// TIA Portal V19 export
DATA_BLOCK "Valves Data"   // DB3
{ S7_Optimized_Access := 'FALSE'; DB_Accessible_From_OPC_UA := 'FALSE' }
// stored: DBAccessibleFromOPCUA false
   VAR RETAIN
      "A/M" : Struct
         R1 : Bool;
         R2 : Bool;
         R3 : Bool;
         R4 : Bool;
         R5 : Bool;
         R6 : Bool;
         R7 : Bool;
         R8 : Bool;
         R9 : Bool;
         R10 : Bool;
         R11 : Bool;
         R12 : Bool;
         R13 : Bool;
         R14 : Bool;
         R15 : Bool;
         R16 : Bool;
         R17 : Bool;
         R18 : Bool;
      END_STRUCT;
      SEMI_AUTO : Struct
         R1 : Bool;
         R2 : Bool;
         R3 : Bool;
         R4 : Bool;
         R5 : Bool;
         R6 : Bool;
         R7 : Bool;
         R8 : Bool;
         R9 : Bool;
         R10 : Bool;
         R11 : Bool;
         R12 : Bool;
         R13 : Bool;
         R14 : Bool;
         R15 : Bool;
         R16 : Bool;
         R17 : Bool;
         R18 : Bool;
      END_STRUCT;
      R1_XV01 : Struct
         MCMD : Bool;
         CMD : Bool;
         RESET : Bool;
         MON_TIME : Time := T#5S;
         STATUS : Int;
         FAULTY : Bool;
      END_STRUCT;
      R1_XV02 : Struct
         MCMD : Bool;
         CMD : Bool;
         RESET : Bool;
         MON_TIME : Time := T#5S;
         STATUS : Int;
         FAULTY : Bool;
      END_STRUCT;
      R1_XV03 : Struct
         MCMD : Bool;
         CMD : Bool;
         RESET : Bool;
         MON_TIME : Time := T#5S;
         STATUS : Int;
         FAULTY : Bool;
      END_STRUCT;
      R1_XV04 : Struct
         MCMD : Bool;
         CMD : Bool;
         RESET : Bool;
         MON_TIME : Time := T#5S;
         STATUS : Int;
         FAULTY : Bool;
      END_STRUCT;
      R1_XV05 : Struct
         MCMD : Bool;
         CMD : Bool;
         RESET : Bool;
         MON_TIME : Time := T#5S;
         STATUS : Int;
         FAULTY : Bool;
      END_STRUCT;
      R1_XV06 : Struct
         MCMD : Bool;
         CMD : Bool;
         RESET : Bool;
         MON_TIME : Time := T#5S;
         STATUS : Int;
         FAULTY : Bool;
      END_STRUCT;
      R1_XV07 : Struct
         MCMD : Bool;
         CMD : Bool;
         RESET : Bool;
         MON_TIME : Time := T#5S;
         STATUS : Int;
         FAULTY : Bool;
      END_STRUCT;
      R1_XV08 : Struct
         MCMD : Bool;
         CMD : Bool;
         RESET : Bool;
         MON_TIME : Time := T#5S;
         STATUS : Int;
         FAULTY : Bool;
      END_STRUCT;
      R1_XV09 : Struct
         MCMD : Bool;
         CMD : Bool;
         RESET : Bool;
         MON_TIME : Time := T#5S;
         STATUS : Int;
         FAULTY : Bool;
      END_STRUCT;
      R1_XV10 : Struct
         MCMD : Bool;
         CMD : Bool;
         RESET : Bool;
         MON_TIME : Time := T#5S;
         STATUS : Int;
         FAULTY : Bool;
      END_STRUCT;
      CCHS_BUXV1501 : Struct
         MCMD : Bool;
         CMD : Bool;
         RESET : Bool;
         MON_TIME : Time := T#5s;
         STATUS : Int;
         FAIL_TO_OPEN : Bool;
         FAIL_TO_CLOSE : Bool;
      END_STRUCT;
      R1_VALVE_FAULT : Struct
         XV01_FAIL_TO_OPEN : Bool;
         XV01_FAIL_TO_CLOSE : Bool;
         XV02_FAIL_TO_OPEN : Bool;
         XV02_FAIL_TO_CLOSE : Bool;
         XV03_FAIL_TO_OPEN : Bool;
         XV03_FAIL_TO_CLOSE : Bool;
         XV04_FAIL_TO_OPEN : Bool;
         XV04_FAIL_TO_CLOSE : Bool;
         XV05_FAIL_TO_OPEN : Bool;
         XV05_FAIL_TO_CLOSE : Bool;
         XV06_FAIL_TO_OPEN : Bool;
         XV06_FAIL_TO_CLOSE : Bool;
         XV07_FAIL_TO_OPEN : Bool;
         XV07_FAIL_TO_CLOSE : Bool;
         XV08_FAIL_TO_OPEN : Bool;
         XV08_FAIL_TO_CLOSE : Bool;
         XV09_FAIL_TO_OPEN : Bool;
         XV09_FAIL_TO_CLOSE : Bool;
         XV010_FAIL_TO_OPEN : Bool;
         XV10_FAIL_TO_CLOSE : Bool;
         CP01_FAIL_TO_RUN : Bool;
         "AG01_FAIL_TO RUN" : Bool;
         CH_CP01_FAIL_TO_RUN : Bool;
         CH_CP02_FAIL_TO_RUN : Bool;
         CH_CP03_FAIL_TO_RUN : Bool;
      END_STRUCT;
      R2_XV01 : Struct
         MCMD : Bool;
         CMD : Bool;
         RESET : Bool;
         MON_TIME : Time := T#5s;
         STATUS : Int;
         FAULTY : Bool;
      END_STRUCT;
      R2_XV02 : Struct
         MCMD : Bool;
         CMD : Bool;
         RESET : Bool;
         MON_TIME : Time := T#5s;
         STATUS : Int;
         FAULTY : Bool;
      END_STRUCT;
      R2_XV03 : Struct
         MCMD : Bool;
         CMD : Bool;
         RESET : Bool;
         MON_TIME : Time := T#5s;
         STATUS : Int;
         FAULTY : Bool;
      END_STRUCT;
      R2_XV04 : Struct
         MCMD : Bool;
         CMD : Bool;
         RESET : Bool;
         MON_TIME : Time := T#5s;
         STATUS : Int;
         FAULTY : Bool;
      END_STRUCT;
      R2_XV05 : Struct
         MCMD : Bool;
         CMD : Bool;
         RESET : Bool;
         MON_TIME : Time := T#5s;
         STATUS : Int;
         FAULTY : Bool;
      END_STRUCT;
      R2_XV06 : Struct
         MCMD : Bool;
         CMD : Bool;
         RESET : Bool;
         MON_TIME : Time := T#5s;
         STATUS : Int;
         FAULTY : Bool;
      END_STRUCT;
      R2_XV07 : Struct
         MCMD : Bool;
         CMD : Bool;
         RESET : Bool;
         MON_TIME : Time := T#5s;
         STATUS : Int;
         FAULTY : Bool;
      END_STRUCT;
      R2_XV08 : Struct
         MCMD : Bool;
         CMD : Bool;
         RESET : Bool;
         MON_TIME : Time := T#5s;
         STATUS : Int;
         FAULTY : Bool;
      END_STRUCT;
      R2_XV09 : Struct
         MCMD : Bool;
         CMD : Bool;
         RESET : Bool;
         MON_TIME : Time := T#5s;
         STATUS : Int;
         FAULTY : Bool;
      END_STRUCT;
      R2_XV10 : Struct
         MCMD : Bool;
         CMD : Bool;
         RESET : Bool;
         MON_TIME : Time := T#5s;
         STATUS : Int;
         FAULTY : Bool;
      END_STRUCT;
      R2_VALVE_FAULT : Struct
         XV01_FAIL_TO_OPEN : Bool;
         XV01_FAIL_TO_CLOSE : Bool;
         XV02_FAIL_TO_OPEN : Bool;
         XV02_FAIL_TO_CLOSE : Bool;
         XV03_FAIL_TO_OPEN : Bool;
         XV03_FAIL_TO_CLOSE : Bool;
         XV04_FAIL_TO_OPEN : Bool;
         XV04_FAIL_TO_CLOSE : Bool;
         XV05_FAIL_TO_OPEN : Bool;
         XV05_FAIL_TO_CLOSE : Bool;
         XV06_FAIL_TO_OPEN : Bool;
         XV06_FAIL_TO_CLOSE : Bool;
         XV07_FAIL_TO_OPEN : Bool;
         XV07_FAIL_TO_CLOSE : Bool;
         XV08_FAIL_TO_OPEN : Bool;
         XV08_FAIL_TO_CLOSE : Bool;
         XV09_FAIL_TO_OPEN : Bool;
         XV09_FAIL_TO_CLOSE : Bool;
         XV010_FAIL_TO_OPEN : Bool;
         XV10_FAIL_TO_CLOSE : Bool;
         CP01_FAIL_TO_RUN : Bool;
         "AG01_FAIL_TO RUN" : Bool;
         CH_CP01_FAIL_TO_RUN : Bool;
         CH_CP02_FAIL_TO_RUN : Bool;
         CH_CP03_FAIL_TO_RUN : Bool;
      END_STRUCT;
      R3_XV01 : Struct
         MCMD : Bool;
         CMD : Bool;
         RESET : Bool;
         MON_TIME : Time := T#5s;
         STATUS : Int;
         FAULTY : Bool;
      END_STRUCT;
      R3_XV02 : Struct
         MCMD : Bool;
         CMD : Bool;
         RESET : Bool;
         MON_TIME : Time := T#5s;
         STATUS : Int;
         FAULTY : Bool;
      END_STRUCT;
      R3_XV03 : Struct
         MCMD : Bool;
         CMD : Bool;
         RESET : Bool;
         MON_TIME : Time := T#5s;
         STATUS : Int;
         FAULTY : Bool;
      END_STRUCT;
      R3_XV04 : Struct
         MCMD : Bool;
         CMD : Bool;
         RESET : Bool;
         MON_TIME : Time := T#5s;
         STATUS : Int;
         FAULTY : Bool;
      END_STRUCT;
      R3_XV05 : Struct
         MCMD : Bool;
         CMD : Bool;
         RESET : Bool;
         MON_TIME : Time := T#5s;
         STATUS : Int;
         FAULTY : Bool;
      END_STRUCT;
      R3_XV06 : Struct
         MCMD : Bool;
         CMD : Bool;
         RESET : Bool;
         MON_TIME : Time := T#5s;
         STATUS : Int;
         FAULTY : Bool;
      END_STRUCT;
      R3_XV07 : Struct
         MCMD : Bool;
         CMD : Bool;
         RESET : Bool;
         MON_TIME : Time := T#5s;
         STATUS : Int;
         FAULTY : Bool;
      END_STRUCT;
      R3_XV08 : Struct
         MCMD : Bool;
         CMD : Bool;
         RESET : Bool;
         MON_TIME : Time := T#5s;
         STATUS : Int;
         FAULTY : Bool;
      END_STRUCT;
      R3_XV09 : Struct
         MCMD : Bool;
         CMD : Bool;
         RESET : Bool;
         MON_TIME : Time := T#5s;
         STATUS : Int;
         FAULTY : Bool;
      END_STRUCT;
      R3_XV10 : Struct
         MCMD : Bool;
         CMD : Bool;
         RESET : Bool;
         MON_TIME : Time := T#5s;
         STATUS : Int;
         FAULTY : Bool;
      END_STRUCT;
      R3_VALVE_FAULT : Struct
         XV01_FAIL_TO_OPEN : Bool;
         XV01_FAIL_TO_CLOSE : Bool;
         XV02_FAIL_TO_OPEN : Bool;
         XV02_FAIL_TO_CLOSE : Bool;
         XV03_FAIL_TO_OPEN : Bool;
         XV03_FAIL_TO_CLOSE : Bool;
         XV04_FAIL_TO_OPEN : Bool;
         XV04_FAIL_TO_CLOSE : Bool;
         XV05_FAIL_TO_OPEN : Bool;
         XV05_FAIL_TO_CLOSE : Bool;
         XV06_FAIL_TO_OPEN : Bool;
         XV06_FAIL_TO_CLOSE : Bool;
         XV07_FAIL_TO_OPEN : Bool;
         XV07_FAIL_TO_CLOSE : Bool;
         XV08_FAIL_TO_OPEN : Bool;
         XV08_FAIL_TO_CLOSE : Bool;
         XV09_FAIL_TO_OPEN : Bool;
         XV09_FAIL_TO_CLOSE : Bool;
         XV010_FAIL_TO_OPEN : Bool;
         XV10_FAIL_TO_CLOSE : Bool;
         CP01_FAIL_TO_RUN : Bool;
         "AG01_FAIL_TO RUN" : Bool;
         CH_CP01_FAIL_TO_RUN : Bool;
         CH_CP02_FAIL_TO_RUN : Bool;
         CH_CP03_FAIL_TO_RUN : Bool;
      END_STRUCT;
      R4_XV01 : Struct
         MCMD : Bool;
         CMD : Bool;
         RESET : Bool;
         MON_TIME : Time := T#5s;
         STATUS : Int;
         FAULTY : Bool;
      END_STRUCT;
      R4_XV02 : Struct
         MCMD : Bool;
         CMD : Bool;
         RESET : Bool;
         MON_TIME : Time := T#5s;
         STATUS : Int;
         FAULTY : Bool;
      END_STRUCT;
      R4_XV03 : Struct
         MCMD : Bool;
         CMD : Bool;
         RESET : Bool;
         MON_TIME : Time := T#5s;
         STATUS : Int;
         FAULTY : Bool;
      END_STRUCT;
      R4_XV04 : Struct
         MCMD : Bool;
         CMD : Bool;
         RESET : Bool;
         MON_TIME : Time := T#5s;
         STATUS : Int;
         FAULTY : Bool;
      END_STRUCT;
      R4_XV05 : Struct
         MCMD : Bool;
         CMD : Bool;
         RESET : Bool;
         MON_TIME : Time := T#5s;
         STATUS : Int;
         FAULTY : Bool;
      END_STRUCT;
      R4_XV06 : Struct
         MCMD : Bool;
         CMD : Bool;
         RESET : Bool;
         MON_TIME : Time := T#5s;
         STATUS : Int;
         FAULTY : Bool;
      END_STRUCT;
      R4_XV07 : Struct
         MCMD : Bool;
         CMD : Bool;
         RESET : Bool;
         MON_TIME : Time := T#5s;
         STATUS : Int;
         FAULTY : Bool;
      END_STRUCT;
      R4_XV08 : Struct
         MCMD : Bool;
         CMD : Bool;
         RESET : Bool;
         MON_TIME : Time := T#5s;
         STATUS : Int;
         FAULTY : Bool;
      END_STRUCT;
      R4_XV09 : Struct
         MCMD : Bool;
         CMD : Bool;
         RESET : Bool;
         MON_TIME : Time := T#5s;
         STATUS : Int;
         FAULTY : Bool;
      END_STRUCT;
      R4_XV10 : Struct
         MCMD : Bool;
         CMD : Bool;
         RESET : Bool;
         MON_TIME : Time := T#5s;
         STATUS : Int;
         FAULTY : Bool;
      END_STRUCT;
      R4_VALVE_FAULT : Struct
         XV01_FAIL_TO_OPEN : Bool;
         XV01_FAIL_TO_CLOSE : Bool;
         XV02_FAIL_TO_OPEN : Bool;
         XV02_FAIL_TO_CLOSE : Bool;
         XV03_FAIL_TO_OPEN : Bool;
         XV03_FAIL_TO_CLOSE : Bool;
         XV04_FAIL_TO_OPEN : Bool;
         XV04_FAIL_TO_CLOSE : Bool;
         XV05_FAIL_TO_OPEN : Bool;
         XV05_FAIL_TO_CLOSE : Bool;
         XV06_FAIL_TO_OPEN : Bool;
         XV06_FAIL_TO_CLOSE : Bool;
         XV07_FAIL_TO_OPEN : Bool;
         XV07_FAIL_TO_CLOSE : Bool;
         XV08_FAIL_TO_OPEN : Bool;
         XV08_FAIL_TO_CLOSE : Bool;
         XV09_FAIL_TO_OPEN : Bool;
         XV09_FAIL_TO_CLOSE : Bool;
         XV010_FAIL_TO_OPEN : Bool;
         XV10_FAIL_TO_CLOSE : Bool;
         CP01_FAIL_TO_RUN : Bool;
         "AG01_FAIL_TO RUN" : Bool;
         CH_CP01_FAIL_TO_RUN : Bool;
         CH_CP02_FAIL_TO_RUN : Bool;
         CH_CP03_FAIL_TO_RUN : Bool;
      END_STRUCT;
      R5_XV01 : Struct
         MCMD : Bool;
         CMD : Bool;
         RESET : Bool;
         MON_TIME : Time := T#5s;
         STATUS : Int;
         FAULTY : Bool;
      END_STRUCT;
      R5_XV02 : Struct
         MCMD : Bool;
         CMD : Bool;
         RESET : Bool;
         MON_TIME : Time := T#5s;
         STATUS : Int;
         FAULTY : Bool;
      END_STRUCT;
      R5_XV03 : Struct
         MCMD : Bool;
         CMD : Bool;
         RESET : Bool;
         MON_TIME : Time := T#5s;
         STATUS : Int;
         FAULTY : Bool;
      END_STRUCT;
      R5_XV04 : Struct
         MCMD : Bool;
         CMD : Bool;
         RESET : Bool;
         MON_TIME : Time := T#5s;
         STATUS : Int;
         FAULTY : Bool;
      END_STRUCT;
      R5_XV05 : Struct
         MCMD : Bool;
         CMD : Bool;
         RESET : Bool;
         MON_TIME : Time := T#5s;
         STATUS : Int;
         FAULTY : Bool;
      END_STRUCT;
      R5_XV06 : Struct
         MCMD : Bool;
         CMD : Bool;
         RESET : Bool;
         MON_TIME : Time := T#5s;
         STATUS : Int;
         FAULTY : Bool;
      END_STRUCT;
      R5_XV07 : Struct
         MCMD : Bool;
         CMD : Bool;
         RESET : Bool;
         MON_TIME : Time := T#5s;
         STATUS : Int;
         FAULTY : Bool;
      END_STRUCT;
      R5_XV08 : Struct
         MCMD : Bool;
         CMD : Bool;
         RESET : Bool;
         MON_TIME : Time := T#5s;
         STATUS : Int;
         FAULTY : Bool;
      END_STRUCT;
      R5_XV09 : Struct
         MCMD : Bool;
         CMD : Bool;
         RESET : Bool;
         MON_TIME : Time := T#5s;
         STATUS : Int;
         FAULTY : Bool;
      END_STRUCT;
      R5_XV10 : Struct
         MCMD : Bool;
         CMD : Bool;
         RESET : Bool;
         MON_TIME : Time := T#5s;
         STATUS : Int;
         FAULTY : Bool;
      END_STRUCT;
      R5_VALVE_FAULT : Struct
         XV01_FAIL_TO_OPEN : Bool;
         XV01_FAIL_TO_CLOSE : Bool;
         XV02_FAIL_TO_OPEN : Bool;
         XV02_FAIL_TO_CLOSE : Bool;
         XV03_FAIL_TO_OPEN : Bool;
         XV03_FAIL_TO_CLOSE : Bool;
         XV04_FAIL_TO_OPEN : Bool;
         XV04_FAIL_TO_CLOSE : Bool;
         XV05_FAIL_TO_OPEN : Bool;
         XV05_FAIL_TO_CLOSE : Bool;
         XV06_FAIL_TO_OPEN : Bool;
         XV06_FAIL_TO_CLOSE : Bool;
         XV07_FAIL_TO_OPEN : Bool;
         XV07_FAIL_TO_CLOSE : Bool;
         XV08_FAIL_TO_OPEN : Bool;
         XV08_FAIL_TO_CLOSE : Bool;
         XV09_FAIL_TO_OPEN : Bool;
         XV09_FAIL_TO_CLOSE : Bool;
         XV010_FAIL_TO_OPEN : Bool;
         XV10_FAIL_TO_CLOSE : Bool;
         CP01_FAIL_TO_RUN : Bool;
         "AG01_FAIL_TO RUN" : Bool;
         CH_CP01_FAIL_TO_RUN : Bool;
         CH_CP02_FAIL_TO_RUN : Bool;
         CH_CP03_FAIL_TO_RUN : Bool;
      END_STRUCT;
      R6_XV01 : Struct
         MCMD : Bool;
         CMD : Bool;
         RESET : Bool;
         MON_TIME : Time := T#5s;
         STATUS : Int;
         FAULTY : Bool;
      END_STRUCT;
      R6_XV02 : Struct
         MCMD : Bool;
         CMD : Bool;
         RESET : Bool;
         MON_TIME : Time := T#5s;
         STATUS : Int;
         FAULTY : Bool;
      END_STRUCT;
      R6_XV03 : Struct
         MCMD : Bool;
         CMD : Bool;
         RESET : Bool;
         MON_TIME : Time := T#5s;
         STATUS : Int;
         FAULTY : Bool;
      END_STRUCT;
      R6_XV04 : Struct
         MCMD : Bool;
         CMD : Bool;
         RESET : Bool;
         MON_TIME : Time := T#5s;
         STATUS : Int;
         FAULTY : Bool;
      END_STRUCT;
      R6_XV05 : Struct
         MCMD : Bool;
         CMD : Bool;
         RESET : Bool;
         MON_TIME : Time := T#5s;
         STATUS : Int;
         FAULTY : Bool;
      END_STRUCT;
      R6_XV06 : Struct
         MCMD : Bool;
         CMD : Bool;
         RESET : Bool;
         MON_TIME : Time := T#5s;
         STATUS : Int;
         FAULTY : Bool;
      END_STRUCT;
      R6_XV07 : Struct
         MCMD : Bool;
         CMD : Bool;
         RESET : Bool;
         MON_TIME : Time := T#5s;
         STATUS : Int;
         FAULTY : Bool;
      END_STRUCT;
      R6_XV08 : Struct
         MCMD : Bool;
         CMD : Bool;
         RESET : Bool;
         MON_TIME : Time := T#5s;
         STATUS : Int;
         FAULTY : Bool;
      END_STRUCT;
      R6_XV09 : Struct
         MCMD : Bool;
         CMD : Bool;
         RESET : Bool;
         MON_TIME : Time := T#5s;
         STATUS : Int;
         FAULTY : Bool;
      END_STRUCT;
      R6_XV10 : Struct
         MCMD : Bool;
         CMD : Bool;
         RESET : Bool;
         MON_TIME : Time := T#5s;
         STATUS : Int;
         FAULTY : Bool;
      END_STRUCT;
      R6_VALVE_FAULT : Struct
         XV01_FAIL_TO_OPEN : Bool;
         XV01_FAIL_TO_CLOSE : Bool;
         XV02_FAIL_TO_OPEN : Bool;
         XV02_FAIL_TO_CLOSE : Bool;
         XV03_FAIL_TO_OPEN : Bool;
         XV03_FAIL_TO_CLOSE : Bool;
         XV04_FAIL_TO_OPEN : Bool;
         XV04_FAIL_TO_CLOSE : Bool;
         XV05_FAIL_TO_OPEN : Bool;
         XV05_FAIL_TO_CLOSE : Bool;
         XV06_FAIL_TO_OPEN : Bool;
         XV06_FAIL_TO_CLOSE : Bool;
         XV07_FAIL_TO_OPEN : Bool;
         XV07_FAIL_TO_CLOSE : Bool;
         XV08_FAIL_TO_OPEN : Bool;
         XV08_FAIL_TO_CLOSE : Bool;
         XV09_FAIL_TO_OPEN : Bool;
         XV09_FAIL_TO_CLOSE : Bool;
         XV010_FAIL_TO_OPEN : Bool;
         XV10_FAIL_TO_CLOSE : Bool;
         CP01_FAIL_TO_RUN : Bool;
         "AG01_FAIL_TO RUN" : Bool;
         CH_CP01_FAIL_TO_RUN : Bool;
         CH_CP02_FAIL_TO_RUN : Bool;
         CH_CP03_FAIL_TO_RUN : Bool;
      END_STRUCT;
      R7_XV01 : Struct
         MCMD : Bool;
         CMD : Bool;
         RESET : Bool;
         MON_TIME : Time := T#5s;
         STATUS : Int;
         FAULTY : Bool;
      END_STRUCT;
      R7_XV02 : Struct
         MCMD : Bool;
         CMD : Bool;
         RESET : Bool;
         MON_TIME : Time := T#5s;
         STATUS : Int;
         FAULTY : Bool;
      END_STRUCT;
      R7_XV03 : Struct
         MCMD : Bool;
         CMD : Bool;
         RESET : Bool;
         MON_TIME : Time := T#5s;
         STATUS : Int;
         FAULTY : Bool;
      END_STRUCT;
      R7_XV04 : Struct
         MCMD : Bool;
         CMD : Bool;
         RESET : Bool;
         MON_TIME : Time := T#5s;
         STATUS : Int;
         FAULTY : Bool;
      END_STRUCT;
      R7_XV05 : Struct
         MCMD : Bool;
         CMD : Bool;
         RESET : Bool;
         MON_TIME : Time := T#5s;
         STATUS : Int;
         FAULTY : Bool;
      END_STRUCT;
      R7_XV06 : Struct
         MCMD : Bool;
         CMD : Bool;
         RESET : Bool;
         MON_TIME : Time := T#5s;
         STATUS : Int;
         FAULTY : Bool;
      END_STRUCT;
      R7_XV07 : Struct
         MCMD : Bool;
         CMD : Bool;
         RESET : Bool;
         MON_TIME : Time := T#5s;
         STATUS : Int;
         FAULTY : Bool;
      END_STRUCT;
      R7_XV08 : Struct
         MCMD : Bool;
         CMD : Bool;
         RESET : Bool;
         MON_TIME : Time := T#5s;
         STATUS : Int;
         FAULTY : Bool;
      END_STRUCT;
      R7_XV09 : Struct
         MCMD : Bool;
         CMD : Bool;
         RESET : Bool;
         MON_TIME : Time := T#5s;
         STATUS : Int;
         FAULTY : Bool;
      END_STRUCT;
      R7_XV10 : Struct
         MCMD : Bool;
         CMD : Bool;
         RESET : Bool;
         MON_TIME : Time := T#5s;
         STATUS : Int;
         FAULTY : Bool;
      END_STRUCT;
      R7_VALVE_FAULT : Struct
         XV01_FAIL_TO_OPEN : Bool;
         XV01_FAIL_TO_CLOSE : Bool;
         XV02_FAIL_TO_OPEN : Bool;
         XV02_FAIL_TO_CLOSE : Bool;
         XV03_FAIL_TO_OPEN : Bool;
         XV03_FAIL_TO_CLOSE : Bool;
         XV04_FAIL_TO_OPEN : Bool;
         XV04_FAIL_TO_CLOSE : Bool;
         XV05_FAIL_TO_OPEN : Bool;
         XV05_FAIL_TO_CLOSE : Bool;
         XV06_FAIL_TO_OPEN : Bool;
         XV06_FAIL_TO_CLOSE : Bool;
         XV07_FAIL_TO_OPEN : Bool;
         XV07_FAIL_TO_CLOSE : Bool;
         XV08_FAIL_TO_OPEN : Bool;
         XV08_FAIL_TO_CLOSE : Bool;
         XV09_FAIL_TO_OPEN : Bool;
         XV09_FAIL_TO_CLOSE : Bool;
         XV010_FAIL_TO_OPEN : Bool;
         XV10_FAIL_TO_CLOSE : Bool;
         CP01_FAIL_TO_RUN : Bool;
         "AG01_FAIL_TO RUN" : Bool;
         CH_CP01_FAIL_TO_RUN : Bool;
         CH_CP02_FAIL_TO_RUN : Bool;
         CH_CP03_FAIL_TO_RUN : Bool;
      END_STRUCT;
      R8_XV01 : Struct
         MCMD : Bool;
         CMD : Bool;
         RESET : Bool;
         MON_TIME : Time := T#5s;
         STATUS : Int;
         FAULTY : Bool;
      END_STRUCT;
      R8_XV02 : Struct
         MCMD : Bool;
         CMD : Bool;
         RESET : Bool;
         MON_TIME : Time := T#5s;
         STATUS : Int;
         FAULTY : Bool;
      END_STRUCT;
      R8_XV03 : Struct
         MCMD : Bool;
         CMD : Bool;
         RESET : Bool;
         MON_TIME : Time := T#5s;
         STATUS : Int;
         FAULTY : Bool;
      END_STRUCT;
      R8_XV04 : Struct
         MCMD : Bool;
         CMD : Bool;
         RESET : Bool;
         MON_TIME : Time := T#5s;
         STATUS : Int;
         FAULTY : Bool;
      END_STRUCT;
      R8_XV05 : Struct
         MCMD : Bool;
         CMD : Bool;
         RESET : Bool;
         MON_TIME : Time := T#5s;
         STATUS : Int;
         FAULTY : Bool;
      END_STRUCT;
      R8_XV06 : Struct
         MCMD : Bool;
         CMD : Bool;
         RESET : Bool;
         MON_TIME : Time := T#5s;
         STATUS : Int;
         FAULTY : Bool;
      END_STRUCT;
      R8_XV07 : Struct
         MCMD : Bool;
         CMD : Bool;
         RESET : Bool;
         MON_TIME : Time := T#5s;
         STATUS : Int;
         FAULTY : Bool;
      END_STRUCT;
      R8_XV08 : Struct
         MCMD : Bool;
         CMD : Bool;
         RESET : Bool;
         MON_TIME : Time := T#5s;
         STATUS : Int;
         FAULTY : Bool;
      END_STRUCT;
      R8_XV09 : Struct
         MCMD : Bool;
         CMD : Bool;
         RESET : Bool;
         MON_TIME : Time := T#5s;
         STATUS : Int;
         FAULTY : Bool;
      END_STRUCT;
      R8_XV10 : Struct
         MCMD : Bool;
         CMD : Bool;
         RESET : Bool;
         MON_TIME : Time := T#5s;
         STATUS : Int;
         FAULTY : Bool;
      END_STRUCT;
      R8_VALVE_FAULT : Struct
         XV01_FAIL_TO_OPEN : Bool;
         XV01_FAIL_TO_CLOSE : Bool;
         XV02_FAIL_TO_OPEN : Bool;
         XV02_FAIL_TO_CLOSE : Bool;
         XV03_FAIL_TO_OPEN : Bool;
         XV03_FAIL_TO_CLOSE : Bool;
         XV04_FAIL_TO_OPEN : Bool;
         XV04_FAIL_TO_CLOSE : Bool;
         XV05_FAIL_TO_OPEN : Bool;
         XV05_FAIL_TO_CLOSE : Bool;
         XV06_FAIL_TO_OPEN : Bool;
         XV06_FAIL_TO_CLOSE : Bool;
         XV07_FAIL_TO_OPEN : Bool;
         XV07_FAIL_TO_CLOSE : Bool;
         XV08_FAIL_TO_OPEN : Bool;
         XV08_FAIL_TO_CLOSE : Bool;
         XV09_FAIL_TO_OPEN : Bool;
         XV09_FAIL_TO_CLOSE : Bool;
         XV010_FAIL_TO_OPEN : Bool;
         XV10_FAIL_TO_CLOSE : Bool;
         CP01_FAIL_TO_RUN : Bool;
         "AG01_FAIL_TO RUN" : Bool;
         CH_CP01_FAIL_TO_RUN : Bool;
         CH_CP02_FAIL_TO_RUN : Bool;
         CH_CP03_FAIL_TO_RUN : Bool;
      END_STRUCT;
      R9_XV01 : Struct
         MCMD : Bool;
         CMD : Bool;
         RESET : Bool;
         MON_TIME : Time := T#5s;
         STATUS : Int;
         FAULTY : Bool;
      END_STRUCT;
      R9_XV02 : Struct
         MCMD : Bool;
         CMD : Bool;
         RESET : Bool;
         MON_TIME : Time := T#5s;
         STATUS : Int;
         FAULTY : Bool;
      END_STRUCT;
      R9_XV03 : Struct
         MCMD : Bool;
         CMD : Bool;
         RESET : Bool;
         MON_TIME : Time := T#5s;
         STATUS : Int;
         FAULTY : Bool;
      END_STRUCT;
      R9_XV04 : Struct
         MCMD : Bool;
         CMD : Bool;
         RESET : Bool;
         MON_TIME : Time := T#5s;
         STATUS : Int;
         FAULTY : Bool;
      END_STRUCT;
      R9_XV05 : Struct
         MCMD : Bool;
         CMD : Bool;
         RESET : Bool;
         MON_TIME : Time := T#5s;
         STATUS : Int;
         FAULTY : Bool;
      END_STRUCT;
      R9_XV06 : Struct
         MCMD : Bool;
         CMD : Bool;
         RESET : Bool;
         MON_TIME : Time := T#5s;
         STATUS : Int;
         FAULTY : Bool;
      END_STRUCT;
      R9_XV07 : Struct
         MCMD : Bool;
         CMD : Bool;
         RESET : Bool;
         MON_TIME : Time := T#5s;
         STATUS : Int;
         FAULTY : Bool;
      END_STRUCT;
      R9_XV08 : Struct
         MCMD : Bool;
         CMD : Bool;
         RESET : Bool;
         MON_TIME : Time := T#5s;
         STATUS : Int;
         FAULTY : Bool;
      END_STRUCT;
      R9_XV09 : Struct
         MCMD : Bool;
         CMD : Bool;
         RESET : Bool;
         MON_TIME : Time := T#5s;
         STATUS : Int;
         FAULTY : Bool;
      END_STRUCT;
      R9_XV10 : Struct
         MCMD : Bool;
         CMD : Bool;
         RESET : Bool;
         MON_TIME : Time := T#5s;
         STATUS : Int;
         FAULTY : Bool;
      END_STRUCT;
      R9_VALVE_FAULT : Struct
         XV01_FAIL_TO_OPEN : Bool;
         XV01_FAIL_TO_CLOSE : Bool;
         XV02_FAIL_TO_OPEN : Bool;
         XV02_FAIL_TO_CLOSE : Bool;
         XV03_FAIL_TO_OPEN : Bool;
         XV03_FAIL_TO_CLOSE : Bool;
         XV04_FAIL_TO_OPEN : Bool;
         XV04_FAIL_TO_CLOSE : Bool;
         XV05_FAIL_TO_OPEN : Bool;
         XV05_FAIL_TO_CLOSE : Bool;
         XV06_FAIL_TO_OPEN : Bool;
         XV06_FAIL_TO_CLOSE : Bool;
         XV07_FAIL_TO_OPEN : Bool;
         XV07_FAIL_TO_CLOSE : Bool;
         XV08_FAIL_TO_OPEN : Bool;
         XV08_FAIL_TO_CLOSE : Bool;
         XV09_FAIL_TO_OPEN : Bool;
         XV09_FAIL_TO_CLOSE : Bool;
         XV010_FAIL_TO_OPEN : Bool;
         XV10_FAIL_TO_CLOSE : Bool;
         CP01_FAIL_TO_RUN : Bool;
         "AG01_FAIL_TO RUN" : Bool;
         CH_CP01_FAIL_TO_RUN : Bool;
         CH_CP02_FAIL_TO_RUN : Bool;
         CH_CP03_FAIL_TO_RUN : Bool;
      END_STRUCT;
      R10_XV01 : Struct
         MCMD : Bool;
         CMD : Bool;
         RESET : Bool;
         MON_TIME : Time := T#5s;
         STATUS : Int;
         FAULTY : Bool;
      END_STRUCT;
      R10_XV02 : Struct
         MCMD : Bool;
         CMD : Bool;
         RESET : Bool;
         MON_TIME : Time := T#5s;
         STATUS : Int;
         FAULTY : Bool;
      END_STRUCT;
      R10_XV03 : Struct
         MCMD : Bool;
         CMD : Bool;
         RESET : Bool;
         MON_TIME : Time := T#5s;
         STATUS : Int;
         FAULTY : Bool;
      END_STRUCT;
      R10_XV04 : Struct
         MCMD : Bool;
         CMD : Bool;
         RESET : Bool;
         MON_TIME : Time := T#5s;
         STATUS : Int;
         FAULTY : Bool;
      END_STRUCT;
      R10_XV05 : Struct
         MCMD : Bool;
         CMD : Bool;
         RESET : Bool;
         MON_TIME : Time := T#5s;
         STATUS : Int;
         FAULTY : Bool;
      END_STRUCT;
      R10_XV06 : Struct
         MCMD : Bool;
         CMD : Bool;
         RESET : Bool;
         MON_TIME : Time := T#5s;
         STATUS : Int;
         FAULTY : Bool;
      END_STRUCT;
      R10_XV07 : Struct
         MCMD : Bool;
         CMD : Bool;
         RESET : Bool;
         MON_TIME : Time := T#5s;
         STATUS : Int;
         FAULTY : Bool;
      END_STRUCT;
      R10_XV08 : Struct
         MCMD : Bool;
         CMD : Bool;
         RESET : Bool;
         MON_TIME : Time := T#5s;
         STATUS : Int;
         FAULTY : Bool;
      END_STRUCT;
      R10_XV09 : Struct
         MCMD : Bool;
         CMD : Bool;
         RESET : Bool;
         MON_TIME : Time := T#5s;
         STATUS : Int;
         FAULTY : Bool;
      END_STRUCT;
      R10_XV10 : Struct
         MCMD : Bool;
         CMD : Bool;
         RESET : Bool;
         MON_TIME : Time := T#5s;
         STATUS : Int;
         FAULTY : Bool;
      END_STRUCT;
      R10_VALVE_FAULT : Struct
         XV01_FAIL_TO_OPEN : Bool;
         XV01_FAIL_TO_CLOSE : Bool;
         XV02_FAIL_TO_OPEN : Bool;
         XV02_FAIL_TO_CLOSE : Bool;
         XV03_FAIL_TO_OPEN : Bool;
         XV03_FAIL_TO_CLOSE : Bool;
         XV04_FAIL_TO_OPEN : Bool;
         XV04_FAIL_TO_CLOSE : Bool;
         XV05_FAIL_TO_OPEN : Bool;
         XV05_FAIL_TO_CLOSE : Bool;
         XV06_FAIL_TO_OPEN : Bool;
         XV06_FAIL_TO_CLOSE : Bool;
         XV07_FAIL_TO_OPEN : Bool;
         XV07_FAIL_TO_CLOSE : Bool;
         XV08_FAIL_TO_OPEN : Bool;
         XV08_FAIL_TO_CLOSE : Bool;
         XV09_FAIL_TO_OPEN : Bool;
         XV09_FAIL_TO_CLOSE : Bool;
         XV010_FAIL_TO_OPEN : Bool;
         XV10_FAIL_TO_CLOSE : Bool;
         CP01_FAIL_TO_RUN : Bool;
         "AG01_FAIL_TO RUN" : Bool;
         CH_CP01_FAIL_TO_RUN : Bool;
         CH_CP02_FAIL_TO_RUN : Bool;
         CH_CP03_FAIL_TO_RUN : Bool;
      END_STRUCT;
      R11_XV01 : Struct
         MCMD : Bool;
         CMD : Bool;
         RESET : Bool;
         MON_TIME : Time := T#5s;
         STATUS : Int;
         FAULTY : Bool;
      END_STRUCT;
      R11_XV02 : Struct
         MCMD : Bool;
         CMD : Bool;
         RESET : Bool;
         MON_TIME : Time := T#5s;
         STATUS : Int;
         FAULTY : Bool;
      END_STRUCT;
      R11_XV03 : Struct
         MCMD : Bool;
         CMD : Bool;
         RESET : Bool;
         MON_TIME : Time := T#5s;
         STATUS : Int;
         FAULTY : Bool;
      END_STRUCT;
      R11_XV04 : Struct
         MCMD : Bool;
         CMD : Bool;
         RESET : Bool;
         MON_TIME : Time := T#5s;
         STATUS : Int;
         FAULTY : Bool;
      END_STRUCT;
      R11_XV05 : Struct
         MCMD : Bool;
         CMD : Bool;
         RESET : Bool;
         MON_TIME : Time := T#5s;
         STATUS : Int;
         FAULTY : Bool;
      END_STRUCT;
      R11_XV06 : Struct
         MCMD : Bool;
         CMD : Bool;
         RESET : Bool;
         MON_TIME : Time := T#5s;
         STATUS : Int;
         FAULTY : Bool;
      END_STRUCT;
      R11_XV07 : Struct
         MCMD : Bool;
         CMD : Bool;
         RESET : Bool;
         MON_TIME : Time := T#5s;
         STATUS : Int;
         FAULTY : Bool;
      END_STRUCT;
      R11_XV08 : Struct
         MCMD : Bool;
         CMD : Bool;
         RESET : Bool;
         MON_TIME : Time := T#5s;
         STATUS : Int;
         FAULTY : Bool;
      END_STRUCT;
      R11_XV09 : Struct
         MCMD : Bool;
         CMD : Bool;
         RESET : Bool;
         MON_TIME : Time := T#5s;
         STATUS : Int;
         FAULTY : Bool;
      END_STRUCT;
      R11_XV10 : Struct
         MCMD : Bool;
         CMD : Bool;
         RESET : Bool;
         MON_TIME : Time := T#5s;
         STATUS : Int;
         FAULTY : Bool;
      END_STRUCT;
      R11_VALVE_FAULT : Struct
         XV01_FAIL_TO_OPEN : Bool;
         XV01_FAIL_TO_CLOSE : Bool;
         XV02_FAIL_TO_OPEN : Bool;
         XV02_FAIL_TO_CLOSE : Bool;
         XV03_FAIL_TO_OPEN : Bool;
         XV03_FAIL_TO_CLOSE : Bool;
         XV04_FAIL_TO_OPEN : Bool;
         XV04_FAIL_TO_CLOSE : Bool;
         XV05_FAIL_TO_OPEN : Bool;
         XV05_FAIL_TO_CLOSE : Bool;
         XV06_FAIL_TO_OPEN : Bool;
         XV06_FAIL_TO_CLOSE : Bool;
         XV07_FAIL_TO_OPEN : Bool;
         XV07_FAIL_TO_CLOSE : Bool;
         XV08_FAIL_TO_OPEN : Bool;
         XV08_FAIL_TO_CLOSE : Bool;
         XV09_FAIL_TO_OPEN : Bool;
         XV09_FAIL_TO_CLOSE : Bool;
         XV010_FAIL_TO_OPEN : Bool;
         XV10_FAIL_TO_CLOSE : Bool;
         CP01_FAIL_TO_RUN : Bool;
         "AG01_FAIL_TO RUN" : Bool;
         CH_CP01_FAIL_TO_RUN : Bool;
         CH_CP02_FAIL_TO_RUN : Bool;
         CH_CP03_FAIL_TO_RUN : Bool;
      END_STRUCT;
      R12_XV01 : Struct
         MCMD : Bool;
         CMD : Bool;
         RESET : Bool;
         MON_TIME : Time := T#5s;
         STATUS : Int;
         FAULTY : Bool;
      END_STRUCT;
      R12_XV02 : Struct
         MCMD : Bool;
         CMD : Bool;
         RESET : Bool;
         MON_TIME : Time := T#5s;
         STATUS : Int;
         FAULTY : Bool;
      END_STRUCT;
      R12_XV03 : Struct
         MCMD : Bool;
         CMD : Bool;
         RESET : Bool;
         MON_TIME : Time := T#5s;
         STATUS : Int;
         FAULTY : Bool;
      END_STRUCT;
      R12_XV04 : Struct
         MCMD : Bool;
         CMD : Bool;
         RESET : Bool;
         MON_TIME : Time := T#5s;
         STATUS : Int;
         FAULTY : Bool;
      END_STRUCT;
      R12_XV05 : Struct
         MCMD : Bool;
         CMD : Bool;
         RESET : Bool;
         MON_TIME : Time := T#5s;
         STATUS : Int;
         FAULTY : Bool;
      END_STRUCT;
      R12_XV06 : Struct
         MCMD : Bool;
         CMD : Bool;
         RESET : Bool;
         MON_TIME : Time := T#5s;
         STATUS : Int;
         FAULTY : Bool;
      END_STRUCT;
      R12_XV07 : Struct
         MCMD : Bool;
         CMD : Bool;
         RESET : Bool;
         MON_TIME : Time := T#5s;
         STATUS : Int;
         FAULTY : Bool;
      END_STRUCT;
      R12_XV08 : Struct
         MCMD : Bool;
         CMD : Bool;
         RESET : Bool;
         MON_TIME : Time := T#5s;
         STATUS : Int;
         FAULTY : Bool;
      END_STRUCT;
      R12_XV09 : Struct
         MCMD : Bool;
         CMD : Bool;
         RESET : Bool;
         MON_TIME : Time := T#5s;
         STATUS : Int;
         FAULTY : Bool;
      END_STRUCT;
      R12_XV10 : Struct
         MCMD : Bool;
         CMD : Bool;
         RESET : Bool;
         MON_TIME : Time := T#5s;
         STATUS : Int;
         FAULTY : Bool;
      END_STRUCT;
      R12_VALVE_FAULT : Struct
         XV01_FAIL_TO_OPEN : Bool;
         XV01_FAIL_TO_CLOSE : Bool;
         XV02_FAIL_TO_OPEN : Bool;
         XV02_FAIL_TO_CLOSE : Bool;
         XV03_FAIL_TO_OPEN : Bool;
         XV03_FAIL_TO_CLOSE : Bool;
         XV04_FAIL_TO_OPEN : Bool;
         XV04_FAIL_TO_CLOSE : Bool;
         XV05_FAIL_TO_OPEN : Bool;
         XV05_FAIL_TO_CLOSE : Bool;
         XV06_FAIL_TO_OPEN : Bool;
         XV06_FAIL_TO_CLOSE : Bool;
         XV07_FAIL_TO_OPEN : Bool;
         XV07_FAIL_TO_CLOSE : Bool;
         XV08_FAIL_TO_OPEN : Bool;
         XV08_FAIL_TO_CLOSE : Bool;
         XV09_FAIL_TO_OPEN : Bool;
         XV09_FAIL_TO_CLOSE : Bool;
         XV010_FAIL_TO_OPEN : Bool;
         XV10_FAIL_TO_CLOSE : Bool;
         CP01_FAIL_TO_RUN : Bool;
         "AG01_FAIL_TO RUN" : Bool;
         CH_CP01_FAIL_TO_RUN : Bool;
         CH_CP02_FAIL_TO_RUN : Bool;
         CH_CP03_FAIL_TO_RUN : Bool;
      END_STRUCT;
      R13_XV01 : Struct
         MCMD : Bool;
         CMD : Bool;
         RESET : Bool;
         MON_TIME : Time := T#5s;
         STATUS : Int;
         FAULTY : Bool;
      END_STRUCT;
      R13_XV02 : Struct
         MCMD : Bool;
         CMD : Bool;
         RESET : Bool;
         MON_TIME : Time := T#5s;
         STATUS : Int;
         FAULTY : Bool;
      END_STRUCT;
      R13_XV03 : Struct
         MCMD : Bool;
         CMD : Bool;
         RESET : Bool;
         MON_TIME : Time := T#5s;
         STATUS : Int;
         FAULTY : Bool;
      END_STRUCT;
      R13_XV04 : Struct
         MCMD : Bool;
         CMD : Bool;
         RESET : Bool;
         MON_TIME : Time := T#5s;
         STATUS : Int;
         FAULTY : Bool;
      END_STRUCT;
      R13_XV05 : Struct
         MCMD : Bool;
         CMD : Bool;
         RESET : Bool;
         MON_TIME : Time := T#5s;
         STATUS : Int;
         FAULTY : Bool;
      END_STRUCT;
      R13_XV06 : Struct
         MCMD : Bool;
         CMD : Bool;
         RESET : Bool;
         MON_TIME : Time := T#5s;
         STATUS : Int;
         FAULTY : Bool;
      END_STRUCT;
      R13_XV07 : Struct
         MCMD : Bool;
         CMD : Bool;
         RESET : Bool;
         MON_TIME : Time := T#5s;
         STATUS : Int;
         FAULTY : Bool;
      END_STRUCT;
      R13_XV08 : Struct
         MCMD : Bool;
         CMD : Bool;
         RESET : Bool;
         MON_TIME : Time := T#5s;
         STATUS : Int;
         FAULTY : Bool;
      END_STRUCT;
      R13_XV09 : Struct
         MCMD : Bool;
         CMD : Bool;
         RESET : Bool;
         MON_TIME : Time := T#5s;
         STATUS : Int;
         FAULTY : Bool;
      END_STRUCT;
      R13_XV10 : Struct
         MCMD : Bool;
         CMD : Bool;
         RESET : Bool;
         MON_TIME : Time := T#5s;
         STATUS : Int;
         FAULTY : Bool;
      END_STRUCT;
      R13_VALVE_FAULT : Struct
         XV01_FAIL_TO_OPEN : Bool;
         XV01_FAIL_TO_CLOSE : Bool;
         XV02_FAIL_TO_OPEN : Bool;
         XV02_FAIL_TO_CLOSE : Bool;
         XV03_FAIL_TO_OPEN : Bool;
         XV03_FAIL_TO_CLOSE : Bool;
         XV04_FAIL_TO_OPEN : Bool;
         XV04_FAIL_TO_CLOSE : Bool;
         XV05_FAIL_TO_OPEN : Bool;
         XV05_FAIL_TO_CLOSE : Bool;
         XV06_FAIL_TO_OPEN : Bool;
         XV06_FAIL_TO_CLOSE : Bool;
         XV07_FAIL_TO_OPEN : Bool;
         XV07_FAIL_TO_CLOSE : Bool;
         XV08_FAIL_TO_OPEN : Bool;
         XV08_FAIL_TO_CLOSE : Bool;
         XV09_FAIL_TO_OPEN : Bool;
         XV09_FAIL_TO_CLOSE : Bool;
         XV010_FAIL_TO_OPEN : Bool;
         XV10_FAIL_TO_CLOSE : Bool;
         CP01_FAIL_TO_RUN : Bool;
         "AG01_FAIL_TO RUN" : Bool;
         CH_CP01_FAIL_TO_RUN : Bool;
         CH_CP02_FAIL_TO_RUN : Bool;
         CH_CP03_FAIL_TO_RUN : Bool;
      END_STRUCT;
      R14_XV01 : Struct
         MCMD : Bool;
         CMD : Bool;
         RESET : Bool;
         MON_TIME : Time := T#5s;
         STATUS : Int;
         FAULTY : Bool;
      END_STRUCT;
      R14_XV02 : Struct
         MCMD : Bool;
         CMD : Bool;
         RESET : Bool;
         MON_TIME : Time := T#5s;
         STATUS : Int;
         FAULTY : Bool;
      END_STRUCT;
      R14_XV03 : Struct
         MCMD : Bool;
         CMD : Bool;
         RESET : Bool;
         MON_TIME : Time := T#5s;
         STATUS : Int;
         FAULTY : Bool;
      END_STRUCT;
      R14_XV04 : Struct
         MCMD : Bool;
         CMD : Bool;
         RESET : Bool;
         MON_TIME : Time := T#5s;
         STATUS : Int;
         FAULTY : Bool;
      END_STRUCT;
      R14_XV05 : Struct
         MCMD : Bool;
         CMD : Bool;
         RESET : Bool;
         MON_TIME : Time := T#5s;
         STATUS : Int;
         FAULTY : Bool;
      END_STRUCT;
      R14_XV06 : Struct
         MCMD : Bool;
         CMD : Bool;
         RESET : Bool;
         MON_TIME : Time := T#5s;
         STATUS : Int;
         FAULTY : Bool;
      END_STRUCT;
      R14_XV07 : Struct
         MCMD : Bool;
         CMD : Bool;
         RESET : Bool;
         MON_TIME : Time := T#5s;
         STATUS : Int;
         FAULTY : Bool;
      END_STRUCT;
      R14_XV08 : Struct
         MCMD : Bool;
         CMD : Bool;
         RESET : Bool;
         MON_TIME : Time := T#5s;
         STATUS : Int;
         FAULTY : Bool;
      END_STRUCT;
      R14_XV09 : Struct
         MCMD : Bool;
         CMD : Bool;
         RESET : Bool;
         MON_TIME : Time := T#5s;
         STATUS : Int;
         FAULTY : Bool;
      END_STRUCT;
      R14_XV10 : Struct
         MCMD : Bool;
         CMD : Bool;
         RESET : Bool;
         MON_TIME : Time := T#5s;
         STATUS : Int;
         FAULTY : Bool;
      END_STRUCT;
      R14_VALVE_FAULT : Struct
         XV01_FAIL_TO_OPEN : Bool;
         XV01_FAIL_TO_CLOSE : Bool;
         XV02_FAIL_TO_OPEN : Bool;
         XV02_FAIL_TO_CLOSE : Bool;
         XV03_FAIL_TO_OPEN : Bool;
         XV03_FAIL_TO_CLOSE : Bool;
         XV04_FAIL_TO_OPEN : Bool;
         XV04_FAIL_TO_CLOSE : Bool;
         XV05_FAIL_TO_OPEN : Bool;
         XV05_FAIL_TO_CLOSE : Bool;
         XV06_FAIL_TO_OPEN : Bool;
         XV06_FAIL_TO_CLOSE : Bool;
         XV07_FAIL_TO_OPEN : Bool;
         XV07_FAIL_TO_CLOSE : Bool;
         XV08_FAIL_TO_OPEN : Bool;
         XV08_FAIL_TO_CLOSE : Bool;
         XV09_FAIL_TO_OPEN : Bool;
         XV09_FAIL_TO_CLOSE : Bool;
         XV010_FAIL_TO_OPEN : Bool;
         XV10_FAIL_TO_CLOSE : Bool;
         CP01_FAIL_TO_RUN : Bool;
         "AG01_FAIL_TO RUN" : Bool;
         CH_CP01_FAIL_TO_RUN : Bool;
         CH_CP02_FAIL_TO_RUN : Bool;
         CH_CP03_FAIL_TO_RUN : Bool;
      END_STRUCT;
      R15_XV01 : Struct
         MCMD : Bool;
         CMD : Bool;
         RESET : Bool;
         MON_TIME : Time := T#5s;
         STATUS : Int;
         FAULTY : Bool;
      END_STRUCT;
      R15_XV02 : Struct
         MCMD : Bool;
         CMD : Bool;
         RESET : Bool;
         MON_TIME : Time := T#5s;
         STATUS : Int;
         FAULTY : Bool;
      END_STRUCT;
      R15_XV03 : Struct
         MCMD : Bool;
         CMD : Bool;
         RESET : Bool;
         MON_TIME : Time := T#5s;
         STATUS : Int;
         FAULTY : Bool;
      END_STRUCT;
      R15_XV04 : Struct
         MCMD : Bool;
         CMD : Bool;
         RESET : Bool;
         MON_TIME : Time := T#5s;
         STATUS : Int;
         FAULTY : Bool;
      END_STRUCT;
      R15_XV05 : Struct
         MCMD : Bool;
         CMD : Bool;
         RESET : Bool;
         MON_TIME : Time := T#5s;
         STATUS : Int;
         FAULTY : Bool;
      END_STRUCT;
      R15_XV06 : Struct
         MCMD : Bool;
         CMD : Bool;
         RESET : Bool;
         MON_TIME : Time := T#5s;
         STATUS : Int;
         FAULTY : Bool;
      END_STRUCT;
      R15_XV07 : Struct
         MCMD : Bool;
         CMD : Bool;
         RESET : Bool;
         MON_TIME : Time := T#5s;
         STATUS : Int;
         FAULTY : Bool;
      END_STRUCT;
      R15_XV08 : Struct
         MCMD : Bool;
         CMD : Bool;
         RESET : Bool;
         MON_TIME : Time := T#5s;
         STATUS : Int;
         FAULTY : Bool;
      END_STRUCT;
      R15_XV09 : Struct
         MCMD : Bool;
         CMD : Bool;
         RESET : Bool;
         MON_TIME : Time := T#5s;
         STATUS : Int;
         FAULTY : Bool;
      END_STRUCT;
      R15_XV10 : Struct
         MCMD : Bool;
         CMD : Bool;
         RESET : Bool;
         MON_TIME : Time := T#5s;
         STATUS : Int;
         FAULTY : Bool;
      END_STRUCT;
      R15_VALVE_FAULT : Struct
         XV01_FAIL_TO_OPEN : Bool;
         XV01_FAIL_TO_CLOSE : Bool;
         XV02_FAIL_TO_OPEN : Bool;
         XV02_FAIL_TO_CLOSE : Bool;
         XV03_FAIL_TO_OPEN : Bool;
         XV03_FAIL_TO_CLOSE : Bool;
         XV04_FAIL_TO_OPEN : Bool;
         XV04_FAIL_TO_CLOSE : Bool;
         XV05_FAIL_TO_OPEN : Bool;
         XV05_FAIL_TO_CLOSE : Bool;
         XV06_FAIL_TO_OPEN : Bool;
         XV06_FAIL_TO_CLOSE : Bool;
         XV07_FAIL_TO_OPEN : Bool;
         XV07_FAIL_TO_CLOSE : Bool;
         XV08_FAIL_TO_OPEN : Bool;
         XV08_FAIL_TO_CLOSE : Bool;
         XV09_FAIL_TO_OPEN : Bool;
         XV09_FAIL_TO_CLOSE : Bool;
         XV010_FAIL_TO_OPEN : Bool;
         XV10_FAIL_TO_CLOSE : Bool;
         CP01_FAIL_TO_RUN : Bool;
         "AG01_FAIL_TO RUN" : Bool;
         CH_CP01_FAIL_TO_RUN : Bool;
         CH_CP02_FAIL_TO_RUN : Bool;
         CH_CP03_FAIL_TO_RUN : Bool;
      END_STRUCT;
      R16_XV01 : Struct
         MCMD : Bool;
         CMD : Bool;
         RESET : Bool;
         MON_TIME : Time := T#5s;
         STATUS : Int;
         FAULTY : Bool;
      END_STRUCT;
      R16_XV02 : Struct
         MCMD : Bool;
         CMD : Bool;
         RESET : Bool;
         MON_TIME : Time := T#5s;
         STATUS : Int;
         FAULTY : Bool;
      END_STRUCT;
      R16_XV03 : Struct
         MCMD : Bool;
         CMD : Bool;
         RESET : Bool;
         MON_TIME : Time := T#5s;
         STATUS : Int;
         FAULTY : Bool;
      END_STRUCT;
      R16_XV04 : Struct
         MCMD : Bool;
         CMD : Bool;
         RESET : Bool;
         MON_TIME : Time := T#5s;
         STATUS : Int;
         FAULTY : Bool;
      END_STRUCT;
      R16_XV05 : Struct
         MCMD : Bool;
         CMD : Bool;
         RESET : Bool;
         MON_TIME : Time := T#5s;
         STATUS : Int;
         FAULTY : Bool;
      END_STRUCT;
      R16_XV06 : Struct
         MCMD : Bool;
         CMD : Bool;
         RESET : Bool;
         MON_TIME : Time := T#5s;
         STATUS : Int;
         FAULTY : Bool;
      END_STRUCT;
      R16_XV07 : Struct
         MCMD : Bool;
         CMD : Bool;
         RESET : Bool;
         MON_TIME : Time := T#5s;
         STATUS : Int;
         FAULTY : Bool;
      END_STRUCT;
      R16_XV08 : Struct
         MCMD : Bool;
         CMD : Bool;
         RESET : Bool;
         MON_TIME : Time := T#5s;
         STATUS : Int;
         FAULTY : Bool;
      END_STRUCT;
      R16_XV09 : Struct
         MCMD : Bool;
         CMD : Bool;
         RESET : Bool;
         MON_TIME : Time := T#5s;
         STATUS : Int;
         FAULTY : Bool;
      END_STRUCT;
      R16_XV10 : Struct
         MCMD : Bool;
         CMD : Bool;
         RESET : Bool;
         MON_TIME : Time := T#5s;
         STATUS : Int;
         FAULTY : Bool;
      END_STRUCT;
      R16_VALVE_FAULT : Struct
         XV01_FAIL_TO_OPEN : Bool;
         XV01_FAIL_TO_CLOSE : Bool;
         XV02_FAIL_TO_OPEN : Bool;
         XV02_FAIL_TO_CLOSE : Bool;
         XV03_FAIL_TO_OPEN : Bool;
         XV03_FAIL_TO_CLOSE : Bool;
         XV04_FAIL_TO_OPEN : Bool;
         XV04_FAIL_TO_CLOSE : Bool;
         XV05_FAIL_TO_OPEN : Bool;
         XV05_FAIL_TO_CLOSE : Bool;
         XV06_FAIL_TO_OPEN : Bool;
         XV06_FAIL_TO_CLOSE : Bool;
         XV07_FAIL_TO_OPEN : Bool;
         XV07_FAIL_TO_CLOSE : Bool;
         XV08_FAIL_TO_OPEN : Bool;
         XV08_FAIL_TO_CLOSE : Bool;
         XV09_FAIL_TO_OPEN : Bool;
         XV09_FAIL_TO_CLOSE : Bool;
         XV010_FAIL_TO_OPEN : Bool;
         XV10_FAIL_TO_CLOSE : Bool;
         CP01_FAIL_TO_RUN : Bool;
         "AG01_FAIL_TO RUN" : Bool;
         CH_CP01_FAIL_TO_RUN : Bool;
         CH_CP02_FAIL_TO_RUN : Bool;
         CH_CP03_FAIL_TO_RUN : Bool;
      END_STRUCT;
      R17_XV01 : Struct
         MCMD : Bool;
         CMD : Bool;
         RESET : Bool;
         MON_TIME : Time := T#5s;
         STATUS : Int;
         FAULTY : Bool;
      END_STRUCT;
      R17_XV02 : Struct
         MCMD : Bool;
         CMD : Bool;
         RESET : Bool;
         MON_TIME : Time := T#5s;
         STATUS : Int;
         FAULTY : Bool;
      END_STRUCT;
      R17_XV03 : Struct
         MCMD : Bool;
         CMD : Bool;
         RESET : Bool;
         MON_TIME : Time := T#5s;
         STATUS : Int;
         FAULTY : Bool;
      END_STRUCT;
      R17_XV04 : Struct
         MCMD : Bool;
         CMD : Bool;
         RESET : Bool;
         MON_TIME : Time := T#5s;
         STATUS : Int;
         FAULTY : Bool;
      END_STRUCT;
      R17_XV05 : Struct
         MCMD : Bool;
         CMD : Bool;
         RESET : Bool;
         MON_TIME : Time := T#5s;
         STATUS : Int;
         FAULTY : Bool;
      END_STRUCT;
      R17_XV06 : Struct
         MCMD : Bool;
         CMD : Bool;
         RESET : Bool;
         MON_TIME : Time := T#5s;
         STATUS : Int;
         FAULTY : Bool;
      END_STRUCT;
      R17_XV07 : Struct
         MCMD : Bool;
         CMD : Bool;
         RESET : Bool;
         MON_TIME : Time := T#5s;
         STATUS : Int;
         FAULTY : Bool;
      END_STRUCT;
      R17_XV08 : Struct
         MCMD : Bool;
         CMD : Bool;
         RESET : Bool;
         MON_TIME : Time := T#5s;
         STATUS : Int;
         FAULTY : Bool;
      END_STRUCT;
      R17_XV09 : Struct
         MCMD : Bool;
         CMD : Bool;
         RESET : Bool;
         MON_TIME : Time := T#5s;
         STATUS : Int;
         FAULTY : Bool;
      END_STRUCT;
      R17_XV10 : Struct
         MCMD : Bool;
         CMD : Bool;
         RESET : Bool;
         MON_TIME : Time := T#5s;
         STATUS : Int;
         FAULTY : Bool;
      END_STRUCT;
      R17_VALVE_FAULT : Struct
         XV01_FAIL_TO_OPEN : Bool;
         XV01_FAIL_TO_CLOSE : Bool;
         XV02_FAIL_TO_OPEN : Bool;
         XV02_FAIL_TO_CLOSE : Bool;
         XV03_FAIL_TO_OPEN : Bool;
         XV03_FAIL_TO_CLOSE : Bool;
         XV04_FAIL_TO_OPEN : Bool;
         XV04_FAIL_TO_CLOSE : Bool;
         XV05_FAIL_TO_OPEN : Bool;
         XV05_FAIL_TO_CLOSE : Bool;
         XV06_FAIL_TO_OPEN : Bool;
         XV06_FAIL_TO_CLOSE : Bool;
         XV07_FAIL_TO_OPEN : Bool;
         XV07_FAIL_TO_CLOSE : Bool;
         XV08_FAIL_TO_OPEN : Bool;
         XV08_FAIL_TO_CLOSE : Bool;
         XV09_FAIL_TO_OPEN : Bool;
         XV09_FAIL_TO_CLOSE : Bool;
         XV010_FAIL_TO_OPEN : Bool;
         XV10_FAIL_TO_CLOSE : Bool;
         CP01_FAIL_TO_RUN : Bool;
         "AG01_FAIL_TO RUN" : Bool;
         CH_CP01_FAIL_TO_RUN : Bool;
         CH_CP02_FAIL_TO_RUN : Bool;
         CH_CP03_FAIL_TO_RUN : Bool;
      END_STRUCT;
      R18_XV01 : Struct
         MCMD : Bool;
         CMD : Bool;
         RESET : Bool;
         MON_TIME : Time := T#5s;
         STATUS : Int;
         FAULTY : Bool;
      END_STRUCT;
      R18_XV02 : Struct
         MCMD : Bool;
         CMD : Bool;
         RESET : Bool;
         MON_TIME : Time := T#5s;
         STATUS : Int;
         FAULTY : Bool;
      END_STRUCT;
      R18_XV03 : Struct
         MCMD : Bool;
         CMD : Bool;
         RESET : Bool;
         MON_TIME : Time := T#5s;
         STATUS : Int;
         FAULTY : Bool;
      END_STRUCT;
      R18_XV04 : Struct
         MCMD : Bool;
         CMD : Bool;
         RESET : Bool;
         MON_TIME : Time := T#5s;
         STATUS : Int;
         FAULTY : Bool;
      END_STRUCT;
      R18_XV05 : Struct
         MCMD : Bool;
         CMD : Bool;
         RESET : Bool;
         MON_TIME : Time := T#5s;
         STATUS : Int;
         FAULTY : Bool;
      END_STRUCT;
      R18_XV06 : Struct
         MCMD : Bool;
         CMD : Bool;
         RESET : Bool;
         MON_TIME : Time := T#5s;
         STATUS : Int;
         FAULTY : Bool;
      END_STRUCT;
      R18_XV07 : Struct
         MCMD : Bool;
         CMD : Bool;
         RESET : Bool;
         MON_TIME : Time := T#5s;
         STATUS : Int;
         FAULTY : Bool;
      END_STRUCT;
      R18_XV08 : Struct
         MCMD : Bool;
         CMD : Bool;
         RESET : Bool;
         MON_TIME : Time := T#5s;
         STATUS : Int;
         FAULTY : Bool;
      END_STRUCT;
      R18_XV09 : Struct
         MCMD : Bool;
         CMD : Bool;
         RESET : Bool;
         MON_TIME : Time := T#5s;
         STATUS : Int;
         FAULTY : Bool;
      END_STRUCT;
      R18_XV10 : Struct
         MCMD : Bool;
         CMD : Bool;
         RESET : Bool;
         MON_TIME : Time := T#5s;
         STATUS : Int;
         FAULTY : Bool;
      END_STRUCT;
      R18_VALVE_FAULT : Struct
         XV01_FAIL_TO_OPEN : Bool;
         XV01_FAIL_TO_CLOSE : Bool;
         XV02_FAIL_TO_OPEN : Bool;
         XV02_FAIL_TO_CLOSE : Bool;
         XV03_FAIL_TO_OPEN : Bool;
         XV03_FAIL_TO_CLOSE : Bool;
         XV04_FAIL_TO_OPEN : Bool;
         XV04_FAIL_TO_CLOSE : Bool;
         XV05_FAIL_TO_OPEN : Bool;
         XV05_FAIL_TO_CLOSE : Bool;
         XV06_FAIL_TO_OPEN : Bool;
         XV06_FAIL_TO_CLOSE : Bool;
         XV07_FAIL_TO_OPEN : Bool;
         XV07_FAIL_TO_CLOSE : Bool;
         XV08_FAIL_TO_OPEN : Bool;
         XV08_FAIL_TO_CLOSE : Bool;
         XV09_FAIL_TO_OPEN : Bool;
         XV09_FAIL_TO_CLOSE : Bool;
         XV010_FAIL_TO_OPEN : Bool;
         XV10_FAIL_TO_CLOSE : Bool;
         CP01_FAIL_TO_RUN : Bool;
         "AG01_FAIL_TO RUN" : Bool;
         CH_CP01_FAIL_TO_RUN : Bool;
         CH_CP02_FAIL_TO_RUN : Bool;
         CH_CP03_FAIL_TO_RUN : Bool;
      END_STRUCT;
      CS_BUXV2001 : Struct
         MCMD : Bool;
         CMD : Bool;
         RESET : Bool;
         MON_TIME : Time := T#5s;
         STATUS : Int;
         FAIL_TO_OPEN : Bool;
         FAIL_TO_CLOSE : Bool;
      END_STRUCT;
      UCHS_BUXV1501 : Struct
         MCMD : Bool;
         CMD : Bool;
         RESET : Bool;
         MON_TIME : Time := T#5s;
         STATUS : Int;
         FAIL_TO_OPEN : Bool;
         FAIL_TO_CLOSE : Bool;
      END_STRUCT;
   END_VAR
BEGIN
END_DATA_BLOCK
